FUNCTION F_BYTES_TO_STRING (* Die ersten SIZE Bytes eines BYTE-Arrays (z. B. von AlPgnRxNew_TP) als STRING auslesen *)
  (* Standard: 61499-1; Description: Copyright (c) 2026 HR Agrartechnik GmbH This program and the accompanying materials are made available under the terms of the Eclipse Public License 2.0 which is available at https://www.eclipse.org/legal/epl-2.0/ SPDX-License-Identifier: EPL-2.0 *)
  (* Version 1.1, 2026-11-14, Franz Höpfinger, HR Agrartechnik GmbH, Eingang LEN in SIZE umbenannt (LEN ist reserviert, Export-Fehler) *)
  (* Version 1.0, 2026-11-13, Franz Höpfinger, HR Agrartechnik GmbH, Initial Version - STRING ueber CAN (mehr als 8 Byte) *)
  PACKAGE logiBUS::utils::dyn_arr;
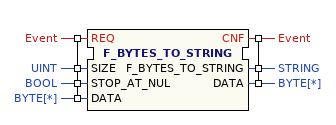
  EVENT_INPUT
    REQ WITH SIZE, STOP_AT_NUL, DATA;
  END_EVENT
  EVENT_OUTPUT
    CNF WITH F_BYTES_TO_STRING, DATA;
  END_EVENT
  VAR_INPUT
    SIZE : UINT; (* Anzahl gueltiger Bytes (z. B. u16DaSize), hoechstens die Groesse von DATA *)
    STOP_AT_NUL : BOOL := TRUE; (* TRUE: Text endet vor dem ersten 16#00 *)
  END_VAR
  VAR_OUTPUT
    F_BYTES_TO_STRING : STRING; (* Text, je Byte 1 Zeichen *)
  END_VAR
  VAR_IN_OUT
    DATA : ARRAY [*] OF BYTE; (* Quellpuffer, z. B. von PROVIDE_ARR_xxxx_BYTE *)
  END_VAR
  BODY IN ST:
PACKAGE logiBUS::utils::dyn_arr;

(* Die ersten SIZE Bytes eines BYTE-Arrays als STRING auslesen *)
FUNCTION F_BYTES_TO_STRING : STRING

VAR_INPUT
	SIZE : UINT; // Anzahl gueltiger Bytes (z. B. u16DaSize)
	STOP_AT_NUL : BOOL := TRUE; // Text endet vor dem ersten 16#00
END_VAR

VAR_IN_OUT
	DATA : ARRAY[*] OF BYTE; // Quellpuffer
END_VAR

VAR_TEMP
	lo : DINT; // erster Index von DATA
	cap : DINT; // Groesse von DATA
	n : DINT; // Anzahl zu lesender Bytes
	i : DINT; // Laufindex
	b : BYTE; // aktuelles Byte
	s : STRING; // Ergebnis in Arbeit
END_VAR

lo := LOWER_BOUND(DATA, 1);
cap := UPPER_BOUND(DATA, 1) - lo + 1;
n := SIZE;
IF n < 0 THEN
	n := 0;
END_IF;
IF n > cap THEN
	n := cap;
END_IF;
s := '';
FOR i := 1 TO n DO
	b := DATA[lo + i - 1];
	IF STOP_AT_NUL AND (b = BYTE#0) THEN
		EXIT;
	END_IF;
	s := CONCAT(s, BYTE_TO_CHAR(b));
END_FOR;
F_BYTES_TO_STRING := s;

END_FUNCTION
  END_BODY
END_FUNCTION
